(* IEC 61131-3 sources: codesys-framework/txt/application/WeVe Visu (library)/Controller/FB_GeneralInputsController, 1 file *)

(* ---- FB_Init.method.st ---- *)
//FB_Init is always available implicitly and it is used primarily for initialization.
//The return value is not evaluated. For a specific influence, you can also declare the
//methods explicitly and provide additional code there with the standard initialization
//code. You can evaluate the return value.
METHOD FB_Init: BOOL
VAR_INPUT
    bInitRetains: BOOL; // TRUE: the retain variables are initialized (reset warm / reset cold)
    bInCopyCode: BOOL;  // TRUE: the instance will be copied to the copy code afterward (online change)

	fbUserRequest 			: I_UserRequestModule;
	fbSignalLamp 			: I_SignalLampModule;
	fbEmergencyStop 		: I_EmergencyStopModule;
END_VAR

// --- BEGIN IMPLEMENTATION ---

_fbUserRequest := fbUserRequest;
_fbSignalLamp := fbSignalLamp;
_fbEmergencyStop := fbEmergencyStop;
